Fanuc KAREL source: kf00115.KL

-- PROVISIONAL review KL for V770-1; original PC SHA256 563cce9e77a4f0a406f08c9b57da304e3ed850ea77336320bd220d4df272598f
-- Incomplete behavior may be omitted. Consult companion uncertainty JSON. Do not deploy.
PROGRAM KF00115
%NOLOCKGROUP
BEGIN
  -- UNRESOLVED_PC offsets 0-1; opcodes 7B
  -- UNRESOLVED_PC offsets 6-18; opcodes 2D,9D,52,7F
  -- UNRESOLVED_PC offsets 23-27; opcodes 7F
  -- UNRESOLVED_PC offsets 32-48; opcodes 27,27,2E,AA,23
  -- UNRESOLVED_PC offsets 53-57; opcodes 7F
END KF00115
